Yaskawa INFORM job: PROG_NA.JBI

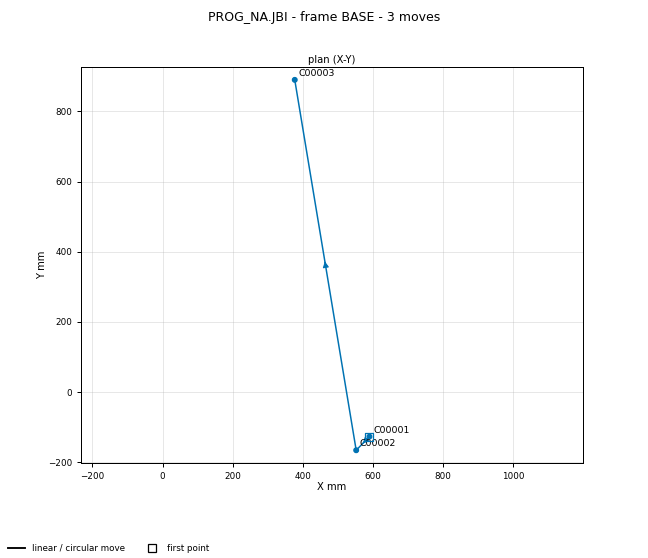
[picture p0: tool path of PROG_NA.JBI in frame BASE, 3 of 5 moves have a stored position in this frame; points joined in program order, loops and branches not executed]
/JOB
//NAME PROG_NA
//POS
///NPOS 5,0,0,0,0,0
///TOOL 9
///POSTYPE PULSE
///PULSE
C00000=10,20,-10,30,-45,60
///TOOL 9
///POSTYPE BASE
///RECTAN
///RCONF 0,0,0,0,0,0,0,0
C00001=589.858,-126.936,665.980,-66.22,8.38,-137.67
C00002=552.056,-165.864,666.221,-67.04,7.80,-141.79
///TOOL 7
C00003=376.936,889.858,655.980,-66.22,8.38,-47.67
///POSTYPE PULSE
///PULSE
C00004=10,20,-10,30,-45,60
//INST
///DATE 2026/10/26 01:19
///COMM Generated using RoboDK
///ATTR SC,RW,RJ
///GROUP1 RB1
NOP
'Program generated by Vertical
'Bot Studio for Motoman GP8 on
' 25/10/2026 12:00:00
'Using nominal kinematics.
'Using Motoman GP8 Base (targe
'ts wrt base):
'0.0,0.0,0.0,0.0,0.0,0.0
'Setting Tool 9 (Spindle):
SETE P00095 (1) 10000
SETE P00095 (2) 0
SETE P00095 (3) 120000
SETE P00095 (4) 0
SETE P00095 (5) 1500
SETE P00095 (6) 0
SETTOOL TL#(9) P00095
MOVJ C00000 VJ=50.00 PL=8
MOVL C00001 V=1000.0 PL=8
MOVL C00002 V=1000.0 PL=0
PAUSE
TIMER T=1.50
MSG "Say "hi" to the operator"
'A long comment line that exce
'eds the usual controller limi
'ts for comments by far, reall
'y
DOUT OT#(12) OFF
DOUT OUT_A ON
WAIT IN#(4)=OFF T=1.00
WAIT IN_B=ON
CALL JOB:PROGRAM
'Using Frame 12 (targets wrt b
'ase):
'250.0,300.0,-10.0,0.0,0.0,90.
'0
'Tool 7 (Tool 7) should be clo
'se to:
'10.0,0.0,120.0,0.0,15.0,0.0
MOVL C00003 V=1000.0 PL=0
MOVJ C00004 VJ=30.00
END
